INTERFACE I_StationManager

METHOD RequestNextStation : I_Station
VAR_INPUT
	CurrentStation : I_Station;
END_VAR
END_METHOD

END_INTERFACE

(* stored: Version 1.1.0.1
   Itf I_StationManager: Id {1c569d71-00c9-4f53-9f61-8233173963d5}
   Method RequestNextStation: Id {d1283a8d-933d-493b-b5bb-6cbad947f201} *)
